(*
SPDX-FileCopyrightText: © 2026 Oleksandr Tiutyk <trofimich@gmail.com>
SPDX-License-Identifier: MIT
License: https://opensource.org/license/mit
*)

(*!
<summary>
Beckhoff EL5101: 1-channel incremental encoder interface terminal (RS422 / TTL, 5 V / 24 V).
</summary>
<description>
Requires enhanced operating mode, available on EL5101 from firmware 14 / hardware 09,
and Standard 32-bit (MDP 511): TxPDO 0x1A04 and RxPDO 0x1603.
Ch1 contains 16-bit status/control and 32-bit counter, latch and preset values.
The normal 16-bit mode and optional frequency/period/timestamp PDOs are outside this model.
When used for I/O, link located fields or their containing buffers to the matching selected PDOs.
The record is not a packed wire buffer; compiler padding is not part of the device specification.
Unlinked/default values do not prove valid I/O. The caller evaluates bus/channel validity before use.
Use one owner task per instance and externally synchronize other access; multi-field snapshots are not atomic.
Copies store data without creating hardware links. Keep borrowed field references valid while consumers are bound.
This passive record performs no validation, synchronization, configuration or protocol advancement.
</description>
*)
TYPE EL5101 :
STRUCT
	Ch1 : INCREMENTAL_ENCODER_CHANNEL;
END_STRUCT
END_TYPE

(* stored: Version 1.1.0.1, ProductVersion 3.1.4026.20
   DUT EL5101: Id {0ba8322e-6441-456d-a430-704be05df22c} *)
